(* IEC 61131-3 sources: model-first-plc-agent-ai/results/T3-W-23, 2 files *)

(* ---- a1_code.st ---- *)
FUNCTION_BLOCK FillingRuntime
VAR_INPUT
    start : BOOL;
    stop : BOOL;
    LSH : BOOL;
    LSHH : BOOL;
    TON_Duration : TIME;
    TOF_Duration : TIME;
END_VAR
VAR_OUTPUT
    fill_valve : BOOL;
    discharge_valve : BOOL;
END_VAR
VAR
    active_state : INT := 0;
    x1 : BOOL;
    ton_q : BOOL;
    tof_q : BOOL;
    filling_timer : TON;
    pause_timer : TOF;
END_VAR

(* Evaluate both timers every scan using the current filling activity. *)
x1 := active_state = 1;

filling_timer(IN := x1, PT := TON_Duration);
pause_timer(IN := x1, PT := TOF_Duration);

ton_q := filling_timer.Q;
tof_q := pause_timer.Q;

(* Execute at most one transition per scan. *)
CASE active_state OF
    0:
        IF start AND NOT stop AND NOT LSH AND NOT LSHH THEN
            active_state := 1;
        END_IF;

    1:
        IF stop OR LSH OR LSHH THEN
            active_state := 0;
        ELSIF ton_q AND NOT stop AND NOT LSH AND NOT LSHH THEN
            active_state := 2;
        END_IF;

    2:
        IF stop OR LSH OR LSHH THEN
            active_state := 0;
        ELSIF NOT tof_q AND NOT stop AND NOT LSH AND NOT LSHH THEN
            active_state := 1;
        END_IF;

ELSE
    active_state := 0;
END_CASE;

(* Continuous, non-stored GRAFCET actions. *)
fill_valve := active_state = 1;
discharge_valve := FALSE;

END_FUNCTION_BLOCK

PROGRAM Main
VAR
    StartCommand AT %IX100.0 : BOOL;
    StopCommand AT %IX100.1 : BOOL;
    LSH AT %IX100.2 : BOOL;
    LSHH AT %IX100.3 : BOOL;
    FillValve AT %QX100.0 : BOOL;
    DischargeValve AT %QX100.1 : BOOL;
END_VAR
VAR
    (* Commissioning defaults; adjust to the required timing parameters. *)
    TON_Duration : TIME := T#5s;
    TOF_Duration : TIME := T#5s;

    start_edge : R_TRIG;
    inputs_initialized : BOOL := FALSE;
    start : BOOL := FALSE;
    runtime_logic : FillingRuntime;
END_VAR

(* Sample the edge detector even on the initialization scan.
   A button already held at startup does not generate a start event. *)
start_edge(CLK := StartCommand);

IF NOT inputs_initialized THEN
    start := FALSE;
    inputs_initialized := TRUE;
ELSE
    start := start_edge.Q;
END_IF;

runtime_logic(
    start := start,
    stop := StopCommand,
    LSH := LSH,
    LSHH := LSHH,
    TON_Duration := TON_Duration,
    TOF_Duration := TOF_Duration
);

FillValve := runtime_logic.fill_valve;
DischargeValve := runtime_logic.discharge_valve;

END_PROGRAM

(* ---- a2_code.st ---- *)
FUNCTION_BLOCK FB_TankFilling
VAR_INPUT
    StartCommand : BOOL;
    StopCommand : BOOL;
    LSH : BOOL;
    LSHH : BOOL;
    TON_Duration : TIME;
    TOF_Duration : TIME;
END_VAR
VAR_OUTPUT
    fill_valve : BOOL;
    discharge_valve : BOOL;
END_VAR
VAR
    sequence_state : INT := 0;
    start_edge : R_TRIG;
    filling_timer : TON;
    pause_timer : TOF;
    start : BOOL;
    stop : BOOL;
    ton_q : BOOL;
    tof_q : BOOL;
    x0 : BOOL;
    x1 : BOOL;
    x2 : BOOL;
END_VAR

start_edge(CLK := StartCommand);
start := start_edge.Q;
stop := StopCommand;

x0 := sequence_state = 0;
x1 := sequence_state = 1;
x2 := sequence_state = 2;

(* Both standard timers measure the activity of the filling step. *)
filling_timer(IN := x1, PT := TON_Duration);
pause_timer(IN := x1, PT := TOF_Duration);

ton_q := filling_timer.Q;
tof_q := pause_timer.Q;

IF stop THEN
    sequence_state := 0;
ELSE
    CASE sequence_state OF
        0:
            IF start AND NOT LSH THEN
                sequence_state := 1;
            END_IF;

        1:
            IF LSH THEN
                sequence_state := 0;
            ELSIF ton_q THEN
                sequence_state := 2;
            END_IF;

        2:
            IF LSH THEN
                sequence_state := 0;
            ELSIF NOT tof_q THEN
                sequence_state := 1;
            END_IF;

        ELSE
            sequence_state := 0;
    END_CASE;
END_IF;

x0 := sequence_state = 0;
x1 := sequence_state = 1;
x2 := sequence_state = 2;

fill_valve := x1;
discharge_valve := FALSE;

END_FUNCTION_BLOCK

PROGRAM Main
VAR
    StartCommand AT %IX100.0 : BOOL;
    StopCommand AT %IX100.1 : BOOL;
    LSH AT %IX100.2 : BOOL;
    LSHH AT %IX100.3 : BOOL;
    FillValve AT %QX100.0 : BOOL;
    DischargeValve AT %QX100.1 : BOOL;
END_VAR
VAR
    tank_controller : FB_TankFilling;
    (* Commissioning defaults; adjust to the required operating durations. *)
    TON_Duration : TIME := T#5s;
    TOF_Duration : TIME := T#5s;
END_VAR

tank_controller(
    StartCommand := StartCommand,
    StopCommand := StopCommand,
    LSH := LSH,
    LSHH := LSHH,
    TON_Duration := TON_Duration,
    TOF_Duration := TOF_Duration
);

FillValve := tank_controller.fill_valve;
DischargeValve := tank_controller.discharge_valve;

END_PROGRAM
